TYPE ET_BOSCH_ManualSetLimits :
(
	eWaitExecute := 0,
	eSetVelo := 5,
	eWfSetVelo := 10,
	eDone := 197,
	eError := 198,
	eNoExecute := 199
);
END_TYPE

(* stored: Version 1.1.0.1, ProductVersion 3.1.4024.15
   DUT ET_BOSCH_ManualSetLimits: Id {50d45081-52da-4bc0-9b39-63fe96bfc4ce} *)
